FUNCTION_BLOCK mF_Mpc
VAR_INPUT
	ssMethodType: SINT;
	flowCurrent: LREAL;
	flowSetpoint: LREAL;
	pressureDifference: LREAL;
END_VAR
VAR_OUTPUT
	valveCommand: LREAL;
END_VAR
VAR
	y_innov: LREAL;
	v: ARRAY[0..1] OF LREAL;
	vseq: ARRAY[0..241] OF LREAL;
	rseq: ARRAY[0..119] OF LREAL;
	a_1: ARRAY[0..243] OF LREAL;
	b: ARRAY[0..243] OF LREAL;
	b_r: ARRAY[0..2] OF LREAL;
	rMin: LREAL;
	b_D: ARRAY[0..8] OF LREAL;
	b_H: ARRAY[0..8] OF LREAL;
	b_U: ARRAY[0..8] OF LREAL;
	cTol: ARRAY[0..243] OF LREAL;
	cTolComputed: BOOL;
	iC: ARRAY[0..243] OF DINT;
	nA: DINT;
	Opt: ARRAY[0..5] OF LREAL;
	Rhs: ARRAY[0..5] OF LREAL;
	DualFeasible: BOOL;
	tmp: DINT;
	ColdReset: BOOL;
	kDrop: DINT;
	Xnorm0: LREAL;
	cMin: LREAL;
	cVal: LREAL;
	z: ARRAY[0..2] OF LREAL;
	t: LREAL;
	iSave: DINT;
	RLinv: ARRAY[0..8] OF LREAL;
	TL: ARRAY[0..8] OF LREAL;
	QQ: ARRAY[0..8] OF LREAL;
	RR: ARRAY[0..8] OF LREAL;
	v_i: DINT;
	k_k: DINT;
	rtb_iAout: ARRAY[0..243] OF BOOL;
	rtb_xest: ARRAY[0..2] OF LREAL;
	i: DINT;
	iC_0: DINT;
	xk: LREAL;
	xk_idx_0: LREAL;
	xk_idx_1: LREAL;
	z_0: LREAL;
	RLinv_tmp: DINT;
	RLinv_tmp_0: DINT;
	rtb_xest_tmp: LREAL;
	exitg1: DINT;
	exitg2: DINT;
	exitg3: DINT;
	exitg4: DINT;
	temp1: BOOL;
	temp2: ARRAY[0..2] OF LREAL;
	temp3: LREAL;
	temp4: ARRAY[0..243] OF LREAL;
	i0_mpcblock_refmd: mpcblock_refmd;
	i0_qr: qr;
	i0_maximum2: maximum2;
	i0_DropConstraint: DropConstraint;
	i0_b_abs: b_abs;
	i0_abs_a: abs_a;
	last_mv_DSTATE: LREAL;
	Memory_PreviousInput: ARRAY[0..243] OF BOOL;
	last_x_PreviousInput: ARRAY[0..2] OF LREAL;
	last_x_InitialCondition: ARRAY[0..2] OF LREAL;
	mF_Mpc_d_a: ARRAY[0..731] OF LREAL := [10.1102866517963, 9.9981210309300046, 9.8827503027042933, 9.7644129935571389, 9.64333938738502, 9.5197517052065965, 9.39386428341519, 9.2658837505365454, 9.1360092024133444, 9.004432375742768, 8.8713378198980148, 8.7369030669692336, 8.601298799963665, 8.4646890191090076, 8.32723120620808, 8.1890764869967949, 8.0503697914612573, 7.9112500120734124, 7.7718501599082854, 7.6322975186091675, 7.4927137961704346, 7.3532152745108172, 7.2139129568129823, 7.0749127126082092, 6.9363154205877446, 6.79821710912512, 6.6607090944962968, 6.5238781167870039, 6.3878064734789888, 6.2525721507092058, 6.1182489521981367, 5.98490662584553, 5.8526109879938435, 5.7214240453615837, 5.5914041146505431, 5.4626059398326934, 5.3350808071241262, 5.2088766576550034, 5.0840381978460005, 4.96060700750311, 4.8386216456440421, 4.7181177540707262, 4.5991281587036212, 4.4816829686946837, 4.3658096733369138, 4.2515332367894159, 4.1388761906378511, 4.0278587243110566, 3.9184987733754468, 3.81081210572957, 3.7048124057219414, 3.6005113562159408, 3.4979187186261744, 3.3970424109513009, 3.29788858382883, 3.2004616946378963, 3.1047645796764534, 3.0107985244397351, 2.9185633320271815, 2.8280573897053647, 2.7392777336547156, 2.6522201119281248, 2.5668790456496784, 2.4832478884819982, 2.4013188843907876, 2.3210832237353118, 2.242531097713631, 2.1656517511914726, 2.0904335339436542, 2.0168639503369952, 1.9449297074836278, 1.8746167618935921, 1.805910364655535, 1.7387951051742592, 1.6732549534937604, 1.6092733012342819, 1.5468330011717719, 1.4859164054879761, 1.4265054027192314, 1.3685814534318335, 1.3121256246516586, 1.2571186230755, 1.2035408270913532, 1.1513723176346458, 1.1005929079071557, 1.0511821719851018, 1.0031194723426136, 0.95638398631651145, 0.910954731538038, 0.86681059035687658, 0.823930333282497, 0.78229264146754784, 0.74187612825770088, 0.70265935983202532, 0.66462087495764166, 0.62773920388206916, 0.591992886386342, 0.55736048902162616, 0.523820621551724, 0.49135195262350245, 0.45993322468693121, 0.42954326818606209, 0.40016101504192586, 0.37176551144796588, 0.34433592999827095, 0.31785158116850964, 0.29229192416911148, 0.26763657718988038, 0.24386532705486785, 0.2209581383059753, 0.19889516173339739, 0.17765674237066328, 0.15722342697167729, 0.137575970986807, 0.11869534505471643, 0.10056274102629219, 0.083159577536662949, 0.066467505140968469, 0.0504684110291919, 0.035144423335029526, -10.1102866517963, -9.9981210309300046, -9.8827503027042933, -9.7644129935571389, -9.64333938738502, -9.5197517052065965, -9.39386428341519, -9.2658837505365454, -9.1360092024133444, -9.004432375742768, -8.8713378198980148, -8.7369030669692336, -8.601298799963665, -8.4646890191090076, -8.32723120620808, -8.1890764869967949, -8.0503697914612573, -7.9112500120734124, -7.7718501599082854, -7.6322975186091675, -7.4927137961704346, -7.3532152745108172, -7.2139129568129823, -7.0749127126082092, -6.9363154205877446, -6.79821710912512, -6.6607090944962968, -6.5238781167870039, -6.3878064734789888, -6.2525721507092058, -6.1182489521981367, -5.98490662584553, -5.8526109879938435, -5.7214240453615837, -5.5914041146505431, -5.4626059398326934, -5.3350808071241262, -5.2088766576550034, -5.0840381978460005, -4.96060700750311, -4.8386216456440421, -4.7181177540707262, -4.5991281587036212, -4.4816829686946837, -4.3658096733369138, -4.2515332367894159, -4.1388761906378511, -4.0278587243110566, -3.9184987733754468, -3.81081210572957, -3.7048124057219414, -3.6005113562159408, -3.4979187186261744, -3.3970424109513009, -3.29788858382883, -3.2004616946378963, -3.1047645796764534, -3.0107985244397351, -2.9185633320271815, -2.8280573897053647, -2.7392777336547156, -2.6522201119281248, -2.5668790456496784, -2.4832478884819982, -2.4013188843907876, -2.3210832237353118, -2.242531097713631, -2.1656517511914726, -2.0904335339436542, -2.0168639503369952, -1.9449297074836278, -1.8746167618935921, -1.805910364655535, -1.7387951051742592, -1.6732549534937604, -1.6092733012342819, -1.5468330011717719, -1.4859164054879761, -1.4265054027192314, -1.3685814534318335, -1.3121256246516586, -1.2571186230755, -1.2035408270913532, -1.1513723176346458, -1.1005929079071557, -1.0511821719851018, -1.0031194723426136, -0.95638398631651145, -0.910954731538038, -0.86681059035687658, -0.823930333282497, -0.78229264146754784, -0.74187612825770088, -0.70265935983202532, -0.66462087495764166, -0.62773920388206916, -0.591992886386342, -0.55736048902162616, -0.523820621551724, -0.49135195262350245, -0.45993322468693121, -0.42954326818606209, -0.40016101504192586, -0.37176551144796588, -0.34433592999827095, -0.31785158116850964, -0.29229192416911148, -0.26763657718988038, -0.24386532705486785, -0.2209581383059753, -0.19889516173339739, -0.17765674237066328, -0.15722342697167729, -0.137575970986807, -0.11869534505471643, -0.10056274102629219, -0.083159577536662949, -0.066467505140968469, -0.0504684110291919, -0.035144423335029526, 0.0, 0.0, 0.0, 0.0, 0.49489060317985373, 0.849211680989655, 1.1869627020934543, 1.5086078890960501, 1.8146039272303969, 2.1053999260864162, 2.3814373892895091, 2.643150191797635, 2.8909645644943867, 3.1252990857639333, 3.3465646797420292, 3.5551646209454835, 3.7514945449905759, 3.9359424651188473, 4.1088887942565426, 4.2707063723416718, 4.4217604986602481, 4.5624089689407183, 4.6930021169629068, 4.8138828604450143, 4.92538675097928, 5.0278420277938505, 5.1215696751252082, 5.2068834829922279, 5.284090111169454, 5.3534891561636471, 5.4153732210039482, 5.470027987662184, 5.5177322919258955, 5.5587582005525915, 5.5933710905395531, 5.6218297303491687, 5.6443863629353537, 5.6612867904220421, 5.6727704602900539, 5.6790705529338288, 5.6804140704545976, 5.677021926561534, 5.6691090374572486, 5.65688441358873, 5.6405512521494554, 5.6203070302228726, 5.5963435984618695, 5.56884727520312, 5.5379989409193433, 5.5039741329166239, 5.4669431401878468, 5.4270710983372, 5.3845180844944194, 5.33943921214112, 5.2919847257750936, 5.2423000953419194, 5.1905261103665827, 5.1367989737210609, 5.0812503949670029, 5.02400768321571, 4.9651938394505954, 4.904927648260232, 4.8433237689328594, 4.780492825865994, 4.7165414982473957, 4.6515726089662159, 4.585685212715628, 4.5189746832506428, 4.451532799767123, 4.3834478323702664, 4.3148046266030011, 4.2456846870068166, 4.1761662596896034, 4.1063244138770107, 4.036231122425737, 3.965955341278975, 3.8955630878460044, 3.8251175182896002, 3.7546790037065736, 3.6843052051883136, 3.6140511477497235, 3.5439692931163842, 3.4741096113611811, 3.404519651382965, 3.3352446102211086, 3.2663274012010461, 3.197808720907072, 3.1297271149798078, 3.0621190427368195, 2.9950189406159184, 2.9284592844416566, 2.8624706505164839, 2.7970817755389228, 2.7323196153519929, 2.668209402525918, 2.6047747027799435, 2.5420374702488178, 2.4800181016002023, 2.4187354890099395, 2.3582070720027279, 2.2984488881663649, 2.2394756227482651, 2.1813006571435007, 2.1239361162841086, 2.067392914939866, 2.0116808029411919, 1.9568084093352314, 1.9027832854865581, 1.8496119471343015, 1.797299915417822, 1.7458517568833669, 1.6952711224844286, 1.6455607855887728, 1.5967226790053528, 1.5487579310445323, 1.5016669006252392, 1.4554492114428432, 1.410103785211708, 1.3656288739965043, 1.3220220916464898, 1.2792804443470613, 1.2374003603029762, 1.1963777185677023, 1.1562078770334181, -0.49489060317985373, -0.849211680989655, -1.1869627020934543, -1.5086078890960501, -1.8146039272303969, -2.1053999260864162, -2.3814373892895091, -2.643150191797635, -2.8909645644943867, -3.1252990857639333, -3.3465646797420292, -3.5551646209454835, -3.7514945449905759, -3.9359424651188473, -4.1088887942565426, -4.2707063723416718, -4.4217604986602481, -4.5624089689407183, -4.6930021169629068, -4.8138828604450143, -4.92538675097928, -5.0278420277938505, -5.1215696751252082, -5.2068834829922279, -5.284090111169454, -5.3534891561636471, -5.4153732210039482, -5.470027987662184, -5.5177322919258955, -5.5587582005525915, -5.5933710905395531, -5.6218297303491687, -5.6443863629353537, -5.6612867904220421, -5.6727704602900539, -5.6790705529338288, -5.6804140704545976, -5.677021926561534, -5.6691090374572486, -5.65688441358873, -5.6405512521494554, -5.6203070302228726, -5.5963435984618695, -5.56884727520312, -5.5379989409193433, -5.5039741329166239, -5.4669431401878468, -5.4270710983372, -5.3845180844944194, -5.33943921214112, -5.2919847257750936, -5.2423000953419194, -5.1905261103665827, -5.1367989737210609, -5.0812503949670029, -5.02400768321571, -4.9651938394505954, -4.904927648260232, -4.8433237689328594, -4.780492825865994, -4.7165414982473957, -4.6515726089662159, -4.585685212715628, -4.5189746832506428, -4.451532799767123, -4.3834478323702664, -4.3148046266030011, -4.2456846870068166, -4.1761662596896034, -4.1063244138770107, -4.036231122425737, -3.965955341278975, -3.8955630878460044, -3.8251175182896002, -3.7546790037065736, -3.6843052051883136, -3.6140511477497235, -3.5439692931163842, -3.4741096113611811, -3.404519651382965, -3.3352446102211086, -3.2663274012010461, -3.197808720907072, -3.1297271149798078, -3.0621190427368195, -2.9950189406159184, -2.9284592844416566, -2.8624706505164839, -2.7970817755389228, -2.7323196153519929, -2.668209402525918, -2.6047747027799435, -2.5420374702488178, -2.4800181016002023, -2.4187354890099395, -2.3582070720027279, -2.2984488881663649, -2.2394756227482651, -2.1813006571435007, -2.1239361162841086, -2.067392914939866, -2.0116808029411919, -1.9568084093352314, -1.9027832854865581, -1.8496119471343015, -1.797299915417822, -1.7458517568833669, -1.6952711224844286, -1.6455607855887728, -1.5967226790053528, -1.5487579310445323, -1.5016669006252392, -1.4554492114428432, -1.410103785211708, -1.3656288739965043, -1.3220220916464898, -1.2792804443470613, -1.2374003603029762, -1.1963777185677023, -1.1562078770334181, 0.0, 0.0, 0.0, 0.0, -1.0, -1.0, -1.0, -1.0, -1.0, -1.0, -1.0, -1.0, -1.0, -1.0, -1.0, -1.0, -1.0, -1.0, -1.0, -1.0, -1.0, -1.0, -1.0, -1.0, -1.0, -1.0, -1.0, -1.0, -1.0, -1.0, -1.0, -1.0, -1.0, -1.0, -1.0, -1.0, -1.0, -1.0, -1.0, -1.0, -1.0, -1.0, -1.0, -1.0, -1.0, -1.0, -1.0, -1.0, -1.0, -1.0, -1.0, -1.0, -1.0, -1.0, -1.0, -1.0, -1.0, -1.0, -1.0, -1.0, -1.0, -1.0, -1.0, -1.0, -1.0, -1.0, -1.0, -1.0, -1.0, -1.0, -1.0, -1.0, -1.0, -1.0, -1.0, -1.0, -1.0, -1.0, -1.0, -1.0, -1.0, -1.0, -1.0, -1.0, -1.0, -1.0, -1.0, -1.0, -1.0, -1.0, -1.0, -1.0, -1.0, -1.0, -1.0, -1.0, -1.0, -1.0, -1.0, -1.0, -1.0, -1.0, -1.0, -1.0, -1.0, -1.0, -1.0, -1.0, -1.0, -1.0, -1.0, -1.0, -1.0, -1.0, -1.0, -1.0, -1.0, -1.0, -1.0, -1.0, -1.0, -1.0, -1.0, -1.0, 1.0, 1.0, 1.0, 1.0, 1.0, 1.0, 1.0, 1.0, 1.0, 1.0, 1.0, 1.0, 1.0, 1.0, 1.0, 1.0, 1.0, 1.0, 1.0, 1.0, 1.0, 1.0, 1.0, 1.0, 1.0, 1.0, 1.0, 1.0, 1.0, 1.0, 1.0, 1.0, 1.0, 1.0, 1.0, 1.0, 1.0, 1.0, 1.0, 1.0, 1.0, 1.0, 1.0, 1.0, 1.0, 1.0, 1.0, 1.0, 1.0, 1.0, 1.0, 1.0, 1.0, 1.0, 1.0, 1.0, 1.0, 1.0, 1.0, 1.0, 1.0, 1.0, 1.0, 1.0, 1.0, 1.0, 1.0, 1.0, 1.0, 1.0, 1.0, 1.0, 1.0, 1.0, 1.0, 1.0, 1.0, 1.0, 1.0, 1.0, 1.0, 1.0, 1.0, 1.0, 1.0, 1.0, 1.0, 1.0, 1.0, 1.0, 1.0, 1.0, 1.0, 1.0, 1.0, 1.0, 1.0, 1.0, 1.0, 1.0, 1.0, 1.0, 1.0, 1.0, 1.0, 1.0, 1.0, 1.0, 1.0, 1.0, 1.0, 1.0, 1.0, 1.0, 1.0, 1.0, 1.0, 1.0, 1.0, 1.0, 0.0, 0.0, 0.0, 0.0];
	mF_Mpc_b_Mlim: ARRAY[0..243] OF LREAL := [0.2, 0.2, 0.2, 0.2, 0.2, 0.2, 0.2, 0.2, 0.2, 0.2, 0.2, 0.2, 0.2, 0.2, 0.2, 0.2, 0.2, 0.2, 0.2, 0.2, 0.2, 0.2, 0.2, 0.2, 0.2, 0.2, 0.2, 0.2, 0.2, 0.2, 0.2, 0.2, 0.2, 0.2, 0.2, 0.2, 0.2, 0.2, 0.2, 0.2, 0.2, 0.2, 0.2, 0.2, 0.2, 0.2, 0.2, 0.2, 0.2, 0.2, 0.2, 0.2, 0.2, 0.2, 0.2, 0.2, 0.2, 0.2, 0.2, 0.2, 0.2, 0.2, 0.2, 0.2, 0.2, 0.2, 0.2, 0.2, 0.2, 0.2, 0.2, 0.2, 0.2, 0.2, 0.2, 0.2, 0.2, 0.2, 0.2, 0.2, 0.2, 0.2, 0.2, 0.2, 0.2, 0.2, 0.2, 0.2, 0.2, 0.2, 0.2, 0.2, 0.2, 0.2, 0.2, 0.2, 0.2, 0.2, 0.2, 0.2, 0.2, 0.2, 0.2, 0.2, 0.2, 0.2, 0.2, 0.2, 0.2, 0.2, 0.2, 0.2, 0.2, 0.2, 0.2, 0.2, 0.2, 0.2, 0.2, 0.2, 0.04, 0.04, 0.04, 0.04, 0.04, 0.04, 0.04, 0.04, 0.04, 0.04, 0.04, 0.04, 0.04, 0.04, 0.04, 0.04, 0.04, 0.04, 0.04, 0.04, 0.04, 0.04, 0.04, 0.04, 0.04, 0.04, 0.04, 0.04, 0.04, 0.04, 0.04, 0.04, 0.04, 0.04, 0.04, 0.04, 0.04, 0.04, 0.04, 0.04, 0.04, 0.04, 0.04, 0.04, 0.04, 0.04, 0.04, 0.04, 0.04, 0.04, 0.04, 0.04, 0.04, 0.04, 0.04, 0.04, 0.04, 0.04, 0.04, 0.04, 0.04, 0.04, 0.04, 0.04, 0.04, 0.04, 0.04, 0.04, 0.04, 0.04, 0.04, 0.04, 0.04, 0.04, 0.04, 0.04, 0.04, 0.04, 0.04, 0.04, 0.04, 0.04, 0.04, 0.04, 0.04, 0.04, 0.04, 0.04, 0.04, 0.04, 0.04, 0.04, 0.04, 0.04, 0.04, 0.04, 0.04, 0.04, 0.04, 0.04, 0.04, 0.04, 0.04, 0.04, 0.04, 0.04, 0.04, 0.04, 0.04, 0.04, 0.04, 0.04, 0.04, 0.04, 0.04, 0.04, 0.04, 0.04, 0.04, 0.04, 1.75, 1.75, -0.25, -0.25];
	mF_Mpc_e_a: ARRAY[0..243] OF LREAL := [-0.00028473180920350741, -0.00064838280152378558, -0.0010871186383875045, -0.0015972149310527575, -0.0021750553811336337, -0.0028171299154482626, -0.0035200328169797839, -0.00428046085366274, -0.0050952114066324721, -0.0059611805995021831, -0.0068753614301614151, -0.0078348419065206853, -0.00883680318755997, -0.0098785177309735454, -0.010957347448640358, -0.012070741871087625, -0.013216236322055611, -0.014391450104213641, -0.015594084697021157, -0.016821921967673122, -0.018072822396016243, -0.019344723314271256, -0.02063563716234695, -0.021943649759483548, -0.023266918592916585, -0.024603671124207489, -0.025952203113843546, -0.027310876964667902, -0.02867812008465969, -0.030052423269545051, -0.031432339105682078, -0.032816480393626085, -0.034203518592746424, -0.035592182287232092, -0.036981255673790715, -0.038369577071313908, -0.039756037452751761, -0.041139578999410086, -0.042519193677855886, -0.043893921839589789, -0.04526285084361819, -0.046625113702033094, -0.047979887748683912, -0.049326393331002638, -0.050663892525022049, -0.051991687873605683, -0.053309121147888459, -0.054615572131907646, -0.055910457430385821, -0.057193229299610078, -0.058463374501335187, -0.05972041317962274, -0.06096389776051344, -0.062193411874415308, -0.063408569301077411, -0.0646090129370057, -0.065794413785165692, -0.066964469966805218, -0.068118905755219825, -0.069257470631273188, -0.070379938360475486, -0.071486106091413787, -0.072575793475319991, -0.073648841806554288, -0.074705113183774638, -0.075744489691556227, -0.076766872602218345, -0.077772181597610637, -0.078760354010605146, -0.079731344086035758, -0.080685122260822376, -0.081621674463012911, -0.082541001429472627, -0.08344311804194729, -0.084328052681223467, -0.085195846599106978, -0.086046553307938353, -0.08688023798736208, -0.087696976908065286, -0.088496856872199881, -0.089279974670201517, -0.090046436553718037, -0.0907963577243595, -0.091529861837982063, -0.092247080524217845, -0.0929481529209633, -0.093633225223539271, -0.094302450248236622, -0.094955987009962314, -0.0955940003137019, -0.096216660359515871, -0.096824142360788817, -0.09741662617545184, -0.0979942959499008, -0.098557339775334651, -0.099105949356240508, -0.099640319690754223, -0.10016064876262748, -0.1006671372445353, -0.10115998821245992, -0.10163940687089022, -0.10210560028857829, -0.10255877714459775, -0.10299914748445149, -0.10342692248597933, -0.10384231423481935, -0.10424553550917975, -0.10463679957368147, -0.10501631998203463, -0.105384310388316, -0.10574098436661702, -0.10608655523883639, -0.10642123591039374, -0.10674523871364502, -0.10705877525878353, -0.1073620562920138, -0.1076552915607895, -0.10793868968590982, -0.10821245804027231, -0.10847680263408387, 0.00028473180920350741, 0.00064838280152378558, 0.0010871186383875045, 0.0015972149310527575, 0.0021750553811336337, 0.0028171299154482626, 0.0035200328169797839, 0.00428046085366274, 0.0050952114066324721, 0.0059611805995021831, 0.0068753614301614151, 0.0078348419065206853, 0.00883680318755997, 0.0098785177309735454, 0.010957347448640358, 0.012070741871087625, 0.013216236322055611, 0.014391450104213641, 0.015594084697021157, 0.016821921967673122, 0.018072822396016243, 0.019344723314271256, 0.02063563716234695, 0.021943649759483548, 0.023266918592916585, 0.024603671124207489, 0.025952203113843546, 0.027310876964667902, 0.02867812008465969, 0.030052423269545051, 0.031432339105682078, 0.032816480393626085, 0.034203518592746424, 0.035592182287232092, 0.036981255673790715, 0.038369577071313908, 0.039756037452751761, 0.041139578999410086, 0.042519193677855886, 0.043893921839589789, 0.04526285084361819, 0.046625113702033094, 0.047979887748683912, 0.049326393331002638, 0.050663892525022049, 0.051991687873605683, 0.053309121147888459, 0.054615572131907646, 0.055910457430385821, 0.057193229299610078, 0.058463374501335187, 0.05972041317962274, 0.06096389776051344, 0.062193411874415308, 0.063408569301077411, 0.0646090129370057, 0.065794413785165692, 0.066964469966805218, 0.068118905755219825, 0.069257470631273188, 0.070379938360475486, 0.071486106091413787, 0.072575793475319991, 0.073648841806554288, 0.074705113183774638, 0.075744489691556227, 0.076766872602218345, 0.077772181597610637, 0.078760354010605146, 0.079731344086035758, 0.080685122260822376, 0.081621674463012911, 0.082541001429472627, 0.08344311804194729, 0.084328052681223467, 0.085195846599106978, 0.086046553307938353, 0.08688023798736208, 0.087696976908065286, 0.088496856872199881, 0.089279974670201517, 0.090046436553718037, 0.0907963577243595, 0.091529861837982063, 0.092247080524217845, 0.0929481529209633, 0.093633225223539271, 0.094302450248236622, 0.094955987009962314, 0.0955940003137019, 0.096216660359515871, 0.096824142360788817, 0.09741662617545184, 0.0979942959499008, 0.098557339775334651, 0.099105949356240508, 0.099640319690754223, 0.10016064876262748, 0.1006671372445353, 0.10115998821245992, 0.10163940687089022, 0.10210560028857829, 0.10255877714459775, 0.10299914748445149, 0.10342692248597933, 0.10384231423481935, 0.10424553550917975, 0.10463679957368147, 0.10501631998203463, 0.105384310388316, 0.10574098436661702, 0.10608655523883639, 0.10642123591039374, 0.10674523871364502, 0.10705877525878353, 0.1073620562920138, 0.1076552915607895, 0.10793868968590982, 0.10821245804027231, 0.10847680263408387, -1.0, -1.0, 1.0, 1.0];
	{attribute 'TcNoSymbol'}
	{attribute 'hide'}
